FUNCTION_BLOCK Fase_Solida (* Fase solida (900): estocagem, alimentacao das prensas C-Press, polimero - HidrycoLib *)
  (* Standard: 61499-2 *)
  (* Version 1.5, 04/11/2026, Hidryco, Hidryco, 1.5: termica das bombas BO-900-01/02/03 NA (cfgTermicaNF = FALSE, campo: ligado = atuada). 1.4: velocidade de partida e PIDs das prensas em Hz (conversao no CLP). 1.3: pidCtl Pid1/2/3 com CycleTime 1000 ms (sem ele o calculo ciclico do pidSC ficava sem periodo). 1.2: sub-CATs Revezamento (horas por soprador, padrao do legado com o nome da elevatoria) e PID (ganho, integral, velocidade minima/maxima das 3 prensas). 1.0: fase solida (900, PCE LODO). Sub-CATs: LIT_900_01/02 (nivel dos tanques, 4-20 mA), FT_900_01/02/03/07 (vazao, comunicacao), SO_900_01/02, BO_900_01..03, BR_900_01/02 (Motor_Generico com ATV), VA_900_01/02, VB_900_03/04, VA_900_06..13 (Valvula_Coester on/off; VA_900_12 futura), AD_900_01..03 (Prensa_Vibropac; AD_900_03 futura), PP_900_01 (Preparador_Vibropac). Campo por symlink ${PATH}: djXXX (disjuntores do PCM LODO, XXX = equipamento), stsEmergenciaPainel (NF), stsMonitTrafo, stsMonitFonte, stsRemota1ComOk, stsRemota2Conexao (INT, connStatusInt); escrita cmdSV01/02/03/04/06/08 (solenoides, manual). *)
  PACKAGE Hidryco.HidrycoLib;
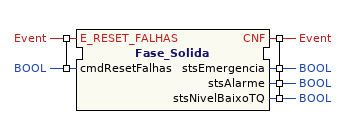
  EVENT_INPUT
    E_RESET_FALHAS WITH cmdResetFalhas; (* Reset pelo processo (fase solida e equipamentos) com cmdResetFalhas = TRUE *)
  END_EVENT
  EVENT_OUTPUT
    CNF WITH stsEmergencia, stsAlarme, stsNivelBaixoTQ; (* Status *)
  END_EVENT
  VAR_INPUT
    cmdResetFalhas : BOOL; (* TRUE = reset (com o evento E_RESET_FALHAS) *)
  END_VAR
  VAR_OUTPUT
    stsEmergencia : BOOL; (* Emergencia do PCM LODO *)
    stsAlarme : BOOL; (* Algum alarme da alimentacao/painel *)
    stsNivelBaixoTQ : BOOL; (* Tanques de estocagem em nivel baixo *)
  END_VAR
  FBS
    IThis : Fase_Solida_HMI(QI := TRUE);
    plcStart1 : plcStart(Prio := 10);
    Tick : E_CYCLE(DT := T#1s);
    Estocagem : basicEstocagemLodo;
    Alimentacao : basicAlimentacaoPrensas;
    Disjuntores1 : SYMLINKMULTIVARDST_854A896E88500D19(QI := TRUE, NAME1 := '$${PATH}djPCE', NAME2 := '$${PATH}djPCM', NAME3 := '$${PATH}djSO01', NAME4 := '$${PATH}djSO02', NAME5 := '$${PATH}djAD01', NAME6 := '$${PATH}djAD02', NAME7 := '$${PATH}djAD03', NAME8 := '$${PATH}djPP01', NAME9 := '$${PATH}djMN01', NAME10 := '$${PATH}djMN02', NAME11 := '$${PATH}djMN03', NAME12 := '$${PATH}djMN04', NAME13 := '$${PATH}djMN05', NAME14 := '$${PATH}djBO01', NAME15 := '$${PATH}djBO02', NAME16 := '$${PATH}djBO03'); {SET_ATTRIBUTE(Configuration.GenericFBType.InterfaceParams, Runtime.System#I:=16;VALUE${I$}:BOOL,BOOL,BOOL,BOOL,BOOL,BOOL,BOOL,BOOL,BOOL,BOOL,BOOL,BOOL,BOOL,BOOL,BOOL,BOOL)}
    Disjuntores2 : SYMLINKMULTIVARDST_854A896E88500D19(QI := TRUE, NAME1 := '$${PATH}djBR01', NAME2 := '$${PATH}djBR02', NAME3 := '$${PATH}djVA01', NAME4 := '$${PATH}djVA02', NAME5 := '$${PATH}djVE01', NAME6 := '$${PATH}djVE02', NAME7 := '$${PATH}djVA06', NAME8 := '$${PATH}djVA07', NAME9 := '$${PATH}djVA08', NAME10 := '$${PATH}djVA09', NAME11 := '$${PATH}djVA10', NAME12 := '$${PATH}djVA11', NAME13 := '$${PATH}djVA12', NAME14 := '$${PATH}djVA13', NAME15 := '$${PATH}djVB03', NAME16 := '$${PATH}djVB04'); {SET_ATTRIBUTE(Configuration.GenericFBType.InterfaceParams, Runtime.System#I:=16;VALUE${I$}:BOOL,BOOL,BOOL,BOOL,BOOL,BOOL,BOOL,BOOL,BOOL,BOOL,BOOL,BOOL,BOOL,BOOL,BOOL,BOOL)}
    Painel : SYMLINKMULTIVARDST_151ACB50A2F8223B2(QI := TRUE, NAME1 := '$${PATH}stsEmergenciaPainel', NAME2 := '$${PATH}stsMonitTrafo', NAME3 := '$${PATH}stsMonitFonte'); {SET_ATTRIBUTE(Configuration.GenericFBType.InterfaceParams, Runtime.System#I:=3;VALUE${I$}:BOOL,BOOL,BOOL)}
    Remota1 : SYMLINKMULTIVARDST_1559B0FF8170C9BA0(QI := TRUE, NAME1 := '$${PATH}stsRemota1ComOk'); {SET_ATTRIBUTE(Configuration.GenericFBType.InterfaceParams, Runtime.System#I:=1;VALUE${I$}:BOOL)}
    Remota2 : SYMLINKMULTIVARDST_5A03F112CD5D470(QI := TRUE, NAME1 := '$${PATH}stsRemota2Conexao'); {SET_ATTRIBUTE(Configuration.GenericFBType.InterfaceParams, Runtime.System#I:=1;VALUE${I$}:INT)}
    Solenoides1 : SYMLINKMULTIVARSRC_151ACB50A2F8223B2(QI := TRUE, NAME1 := '$${PATH}cmdSV01', NAME2 := '$${PATH}cmdSV02', NAME3 := '$${PATH}cmdSV03'); {SET_ATTRIBUTE(Configuration.GenericFBType.InterfaceParams, Runtime.System#I:=3;VALUE${I$}:BOOL,BOOL,BOOL)}
    Solenoides2 : SYMLINKMULTIVARSRC_151ACB50A2F8223B2(QI := TRUE, NAME1 := '$${PATH}cmdSV04', NAME2 := '$${PATH}cmdSV06', NAME3 := '$${PATH}cmdSV08'); {SET_ATTRIBUTE(Configuration.GenericFBType.InterfaceParams, Runtime.System#I:=3;VALUE${I$}:BOOL,BOOL,BOOL)}
    PersBO1 : PERSISTENCE_20652AC5DB8BA8AD5(QI := TRUE); {SET_ATTRIBUTE(Configuration.GenericFBType.InterfaceParams, Runtime.Standard#I:=3;input${I$}:UINT,UINT,UDINT)}
    PersBO2 : PERSISTENCE_20652AC5DB8BA8AD5(QI := TRUE); {SET_ATTRIBUTE(Configuration.GenericFBType.InterfaceParams, Runtime.Standard#I:=3;input${I$}:UINT,UINT,UDINT)}
    PersBO3 : PERSISTENCE_20652AC5DB8BA8AD5(QI := TRUE); {SET_ATTRIBUTE(Configuration.GenericFBType.InterfaceParams, Runtime.Standard#I:=3;input${I$}:UINT,UINT,UDINT)}
    Pid1 : pidCtl(CycleTime := 1000, Direction := TRUE, Bump := FALSE, ProhibitOutInc := FALSE, ProhibitOutDec := FALSE);
    Pid2 : pidCtl(CycleTime := 1000, Direction := TRUE, Bump := FALSE, ProhibitOutInc := FALSE, ProhibitOutDec := FALSE);
    Pid3 : pidCtl(CycleTime := 1000, Direction := TRUE, Bump := FALSE, ProhibitOutInc := FALSE, ProhibitOutDec := FALSE);
    LIT_900_01 : Sensor_Generico(pin_FC98F78ABCBC0A7E := TRUE, pin_CC8EEC06FF0C4430 := 'm', pin_6D3A2524C5D0F0D1 := 2);
    LIT_900_02 : Sensor_Generico(pin_FC98F78ABCBC0A7E := TRUE, pin_CC8EEC06FF0C4430 := 'm', pin_6D3A2524C5D0F0D1 := 2);
    FT_900_01 : Sensor_Generico(pin_D46B37D45FD5AF5D := TRUE, pin_0ECE7B3867B02E0B := TRUE, pin_CC8EEC06FF0C4430 := 'm3/h', pin_6D3A2524C5D0F0D1 := 1);
    FT_900_02 : Sensor_Generico(pin_D46B37D45FD5AF5D := TRUE, pin_0ECE7B3867B02E0B := TRUE, pin_CC8EEC06FF0C4430 := 'm3/h', pin_6D3A2524C5D0F0D1 := 1);
    FT_900_03 : Sensor_Generico(pin_D46B37D45FD5AF5D := TRUE, pin_0ECE7B3867B02E0B := TRUE, pin_CC8EEC06FF0C4430 := 'm3/h', pin_6D3A2524C5D0F0D1 := 1);
    FT_900_07 : Sensor_Generico(pin_D46B37D45FD5AF5D := TRUE, pin_0ECE7B3867B02E0B := TRUE, pin_CC8EEC06FF0C4430 := 'm3/h', pin_6D3A2524C5D0F0D1 := 1);
    SO_900_01 : Motor_Generico(pin_63EFEFB7C85EC93E := TRUE, pin_39489193B7758574 := 600.0);
    SO_900_02 : Motor_Generico(pin_63EFEFB7C85EC93E := TRUE, pin_39489193B7758574 := 600.0);
    BO_900_01 : Motor_Generico(pin_63EFEFB7C85EC93E := TRUE, pin_39489193B7758574 := 600.0, pin_66763E13F70A4420 := FALSE);
    BO_900_02 : Motor_Generico(pin_63EFEFB7C85EC93E := TRUE, pin_39489193B7758574 := 600.0, pin_66763E13F70A4420 := FALSE);
    BO_900_03 : Motor_Generico(pin_63EFEFB7C85EC93E := TRUE, pin_39489193B7758574 := 600.0, pin_66763E13F70A4420 := FALSE);
    BR_900_01 : Motor_Generico(pin_63EFEFB7C85EC93E := TRUE, pin_39489193B7758574 := 600.0);
    BR_900_02 : Motor_Generico(pin_63EFEFB7C85EC93E := TRUE, pin_39489193B7758574 := 600.0);
    VA_900_01 : Atuador_Coester;
    VA_900_02 : Atuador_Coester;
    VB_900_03 : Atuador_Coester;
    VB_900_04 : Atuador_Coester;
    VA_900_06 : Atuador_Coester;
    VA_900_07 : Atuador_Coester;
    VA_900_08 : Atuador_Coester;
    VA_900_09 : Atuador_Coester;
    VA_900_10 : Atuador_Coester;
    VA_900_11 : Atuador_Coester;
    VA_900_12 : Atuador_Coester(pin_FFAFC48D6FD3FF02 := FALSE);
    VA_900_13 : Atuador_Coester;
    AD_900_01 : Prensa_Vibropac;
    AD_900_02 : Prensa_Vibropac;
    AD_900_03 : Prensa_Vibropac(pin_FF2D8D14693482D2 := FALSE);
    PP_900_01 : Preparador_Vibropac;
    AlarmeSopradores : ALARM_BIT(TYPE := 1, ACKTYPE_1 := 2, ACTIVE := TRUE); {SET_ATTRIBUTE(HMI.AlarmText, Tanques de lodo: nenhum soprador disponível)}
    AlarmeNivelTQ : ALARM_BIT(TYPE := 1, ACKTYPE_1 := 2, ACTIVE := TRUE); {SET_ATTRIBUTE(HMI.AlarmText, Tanques de lodo: nível baixo - bombas suspensas)} {SET_ATTRIBUTE(HMI.AlarmClass, Warning)}
    AlarmeEmergencia : ALARM_BIT(TYPE := 1, ACKTYPE_1 := 2, ACTIVE := TRUE); {SET_ATTRIBUTE(HMI.AlarmText, PCM LODO: emergência acionada)}
    AlarmeRemota : ALARM_BIT(TYPE := 1, ACKTYPE_1 := 2, ACTIVE := TRUE); {SET_ATTRIBUTE(HMI.AlarmText, PCE LODO: remota sem comunicação)} {SET_ATTRIBUTE(HMI.AlarmClass, Warning)}
    AlarmeDisjuntor : ALARM_BIT(TYPE := 1, ACKTYPE_1 := 2, ACTIVE := TRUE); {SET_ATTRIBUTE(HMI.AlarmText, PCM LODO: disjuntor desligado)} {SET_ATTRIBUTE(HMI.AlarmClass, Warning)}
    AlarmeRota : ALARM_BIT(TYPE := 1, ACKTYPE_1 := 2, ACTIVE := TRUE); {SET_ATTRIBUTE(HMI.AlarmText, Alimentação das prensas: válvulas da rota não abriram)}
    AlarmeSemBomba : ALARM_BIT(TYPE := 1, ACKTYPE_1 := 2, ACTIVE := TRUE); {SET_ATTRIBUTE(HMI.AlarmText, Alimentação das prensas: sem bomba disponível)} {SET_ATTRIBUTE(HMI.AlarmClass, Warning)}
    AlarmeSemPartir : ALARM_BIT(TYPE := 1, ACKTYPE_1 := 2, ACTIVE := TRUE); {SET_ATTRIBUTE(HMI.AlarmText, Alimentação das prensas: prensa não partiu)} {SET_ATTRIBUTE(HMI.AlarmClass, Warning)}
    AlarmeFT : ALARM_BIT(TYPE := 1, ACKTYPE_1 := 2, ACTIVE := TRUE); {SET_ATTRIBUTE(HMI.AlarmText, Alimentação das prensas: medidor de vazão em falha)} {SET_ATTRIBUTE(HMI.AlarmClass, Warning)}
    Revezamento : Controle_Revezamento_2;
    PID : Controle_PID;
  END_FBS
  EVENT_CONNECTIONS
    plcStart1.FIRST_INIT TO IThis.F45AEED5C0881751;
    plcStart1.REDO_INIT TO IThis.F45AEED5C0881751;
    IThis.89CE2E9FA670B6C6 TO Disjuntores1.INIT;
    Disjuntores1.INITO TO Disjuntores2.INIT;
    Disjuntores2.INITO TO Painel.INIT;
    Painel.INITO TO Remota1.INIT;
    Remota1.INITO TO Remota2.INIT;
    Remota2.INITO TO Solenoides1.INIT;
    Solenoides1.INITO TO Solenoides2.INIT;
    Solenoides2.INITO TO Estocagem.243DC77CA0D0953F;
    Estocagem.5F76B62564497316 TO Alimentacao.13FEA6D5249A7B77;
    Alimentacao.8D3D86F80598A7BB TO IThis.AD1CFD9CF87E7BE8;
    Alimentacao.8D3D86F80598A7BB TO Tick.START;
    Alimentacao.8D3D86F80598A7BB TO PersBO1.INIT;
    PersBO1.INITO TO PersBO1.READ;
    PersBO1.READCNF TO Alimentacao.08CA7CB6A8F97690;
    Alimentacao.557985467D809489 TO PersBO1.WRITE;
    PersBO1.INITO TO PersBO2.INIT;
    PersBO2.INITO TO PersBO2.READ;
    PersBO2.READCNF TO Alimentacao.08CA7CB6A8F97690;
    Alimentacao.557985467D809489 TO PersBO2.WRITE;
    PersBO2.INITO TO PersBO3.INIT;
    PersBO3.INITO TO PersBO3.READ;
    PersBO3.READCNF TO Alimentacao.08CA7CB6A8F97690;
    Alimentacao.557985467D809489 TO PersBO3.WRITE;
    PersBO3.INITO TO AlarmeSopradores.INIT;
    AlarmeSopradores.INITO TO AlarmeSopradores.REQ_INITDATA;
    AlarmeSopradores.CNF_INITDATA TO AlarmeSopradores.ACTIVATE;
    AlarmeNivelTQ.INITO TO AlarmeNivelTQ.REQ_INITDATA;
    AlarmeNivelTQ.CNF_INITDATA TO AlarmeNivelTQ.ACTIVATE;
    AlarmeSopradores.INITO TO AlarmeNivelTQ.INIT;
    AlarmeEmergencia.INITO TO AlarmeEmergencia.REQ_INITDATA;
    AlarmeEmergencia.CNF_INITDATA TO AlarmeEmergencia.ACTIVATE;
    AlarmeNivelTQ.INITO TO AlarmeEmergencia.INIT;
    AlarmeRemota.INITO TO AlarmeRemota.REQ_INITDATA;
    AlarmeRemota.CNF_INITDATA TO AlarmeRemota.ACTIVATE;
    AlarmeEmergencia.INITO TO AlarmeRemota.INIT;
    AlarmeDisjuntor.INITO TO AlarmeDisjuntor.REQ_INITDATA;
    AlarmeDisjuntor.CNF_INITDATA TO AlarmeDisjuntor.ACTIVATE;
    AlarmeRemota.INITO TO AlarmeDisjuntor.INIT;
    AlarmeRota.INITO TO AlarmeRota.REQ_INITDATA;
    AlarmeRota.CNF_INITDATA TO AlarmeRota.ACTIVATE;
    AlarmeDisjuntor.INITO TO AlarmeRota.INIT;
    AlarmeSemBomba.INITO TO AlarmeSemBomba.REQ_INITDATA;
    AlarmeSemBomba.CNF_INITDATA TO AlarmeSemBomba.ACTIVATE;
    AlarmeRota.INITO TO AlarmeSemBomba.INIT;
    AlarmeSemPartir.INITO TO AlarmeSemPartir.REQ_INITDATA;
    AlarmeSemPartir.CNF_INITDATA TO AlarmeSemPartir.ACTIVATE;
    AlarmeSemBomba.INITO TO AlarmeSemPartir.INIT;
    AlarmeFT.INITO TO AlarmeFT.REQ_INITDATA;
    AlarmeFT.CNF_INITDATA TO AlarmeFT.ACTIVATE;
    AlarmeSemPartir.INITO TO AlarmeFT.INIT;
    AlarmeFT.INITO TO plcStart1.ACK_FIRST;
    Tick.EO TO Estocagem.E8C8FA9D941AAB25;
    Tick.EO TO Alimentacao.97FA92419A632264;
    Disjuntores1.CNF TO Alimentacao.856DAE0A3F3D97F7;
    Disjuntores2.CNF TO Alimentacao.856DAE0A3F3D97F7;
    Painel.CNF TO Alimentacao.19B51840153EBC5A;
    Remota1.CNF TO Alimentacao.939B3751BD07756D;
    Remota2.CNF TO Alimentacao.5748134B24BEF763;
    SO_900_01.9D4F26EE27EDF5B9 TO Estocagem.DFFA20E8FEFD328B;
    Estocagem.A37D04399243417C TO SO_900_01.21070E4B73BFECDC;
    SO_900_02.9D4F26EE27EDF5B9 TO Estocagem.DFFA20E8FEFD328B;
    Estocagem.A37D04399243417C TO SO_900_02.21070E4B73BFECDC;
    LIT_900_01.28A380156DB271B8 TO Estocagem.EA4444D55C79B643;
    LIT_900_02.28A380156DB271B8 TO Estocagem.EA4444D55C79B643;
    Alimentacao.8A05961272844DF6 TO Estocagem.EBAA94C91027AB04;
    Estocagem.820328527C60D44B TO VA_900_01.6AE7937B5439A162;
    Estocagem.820328527C60D44B TO VA_900_02.6AE7937B5439A162;
    Estocagem.820328527C60D44B TO VB_900_03.6AE7937B5439A162;
    Estocagem.820328527C60D44B TO VB_900_04.6AE7937B5439A162;
    Estocagem.DD4EDADF061294FF TO Alimentacao.CBCF1D50DEE68A86;
    AD_900_01.8111B44229D619D2 TO Alimentacao.38F5F6E182F651D4;
    Alimentacao.9C532436C7A3B461 TO AD_900_01.7E5F12997195C3C2;
    AD_900_02.8111B44229D619D2 TO Alimentacao.38F5F6E182F651D4;
    Alimentacao.9C532436C7A3B461 TO AD_900_02.7E5F12997195C3C2;
    AD_900_03.8111B44229D619D2 TO Alimentacao.38F5F6E182F651D4;
    Alimentacao.9C532436C7A3B461 TO AD_900_03.7E5F12997195C3C2;
    BO_900_01.9D4F26EE27EDF5B9 TO Alimentacao.CA246CEBE60B1023;
    Alimentacao.7490FED3332AEC1E TO BO_900_01.21070E4B73BFECDC;
    BO_900_02.9D4F26EE27EDF5B9 TO Alimentacao.CA246CEBE60B1023;
    Alimentacao.7490FED3332AEC1E TO BO_900_02.21070E4B73BFECDC;
    BO_900_03.9D4F26EE27EDF5B9 TO Alimentacao.CA246CEBE60B1023;
    Alimentacao.7490FED3332AEC1E TO BO_900_03.21070E4B73BFECDC;
    Alimentacao.7490FED3332AEC1E TO BR_900_01.21070E4B73BFECDC;
    Alimentacao.7490FED3332AEC1E TO BR_900_02.21070E4B73BFECDC;
    VA_900_06.CF6616D3CB5312F6 TO Alimentacao.6647071B86B2ADCE;
    Alimentacao.B985DE359C566AD4 TO VA_900_06.6AE7937B5439A162;
    VA_900_07.CF6616D3CB5312F6 TO Alimentacao.6647071B86B2ADCE;
    Alimentacao.B985DE359C566AD4 TO VA_900_07.6AE7937B5439A162;
    VA_900_08.CF6616D3CB5312F6 TO Alimentacao.6647071B86B2ADCE;
    Alimentacao.B985DE359C566AD4 TO VA_900_08.6AE7937B5439A162;
    VA_900_09.CF6616D3CB5312F6 TO Alimentacao.6647071B86B2ADCE;
    Alimentacao.B985DE359C566AD4 TO VA_900_09.6AE7937B5439A162;
    VA_900_10.CF6616D3CB5312F6 TO Alimentacao.6647071B86B2ADCE;
    Alimentacao.B985DE359C566AD4 TO VA_900_10.6AE7937B5439A162;
    VA_900_11.CF6616D3CB5312F6 TO Alimentacao.6647071B86B2ADCE;
    Alimentacao.B985DE359C566AD4 TO VA_900_11.6AE7937B5439A162;
    VA_900_12.CF6616D3CB5312F6 TO Alimentacao.6647071B86B2ADCE;
    Alimentacao.B985DE359C566AD4 TO VA_900_12.6AE7937B5439A162;
    VA_900_13.CF6616D3CB5312F6 TO Alimentacao.6647071B86B2ADCE;
    Alimentacao.B985DE359C566AD4 TO VA_900_13.6AE7937B5439A162;
    FT_900_01.28A380156DB271B8 TO Alimentacao.48ABB9D9BB2D6CEE;
    IThis.2286FBFA7E7E3034 TO Pid1.REQ_SP;
    FT_900_01.28A380156DB271B8 TO Pid1.REQ;
    Alimentacao.CF7635F428763261 TO Pid1.REQ;
    Pid1.CNF TO Alimentacao.37F5128277E33C7D;
    Pid1.C_CNF TO Alimentacao.37F5128277E33C7D;
    FT_900_02.28A380156DB271B8 TO Alimentacao.48ABB9D9BB2D6CEE;
    IThis.2286FBFA7E7E3034 TO Pid2.REQ_SP;
    FT_900_02.28A380156DB271B8 TO Pid2.REQ;
    Alimentacao.CF7635F428763261 TO Pid2.REQ;
    Pid2.CNF TO Alimentacao.37F5128277E33C7D;
    Pid2.C_CNF TO Alimentacao.37F5128277E33C7D;
    FT_900_03.28A380156DB271B8 TO Alimentacao.48ABB9D9BB2D6CEE;
    IThis.2286FBFA7E7E3034 TO Pid3.REQ_SP;
    FT_900_03.28A380156DB271B8 TO Pid3.REQ;
    Alimentacao.CF7635F428763261 TO Pid3.REQ;
    Pid3.CNF TO Alimentacao.37F5128277E33C7D;
    Pid3.C_CNF TO Alimentacao.37F5128277E33C7D;
    PP_900_01.0264E737EBBCA257 TO Alimentacao.2E29057D22A77FC3;
    Alimentacao.FAFF2EF1C05DA77F TO PP_900_01.8E41CA7EF16C6739;
    Alimentacao.F922E54EB08BF260 TO Solenoides1.REQ;
    Alimentacao.F922E54EB08BF260 TO Solenoides2.REQ;
    IThis.2286FBFA7E7E3034 TO Estocagem.C2DAB560DFFB8D5C;
    IThis.2286FBFA7E7E3034 TO Alimentacao.912D39602F9C91C5;
    IThis.94340A1957F06E33 TO Alimentacao.477B3CB066C0064B;
    IThis.DA6F3DD5304C4EDD TO Alimentacao.B672F1361E424ACE;
    IThis.EA322A066409681E TO Alimentacao.FBC24ECA7AD15CA0;
    Estocagem.12E6850BBBD0B68E TO IThis.0FDAAD8F71C680CA;
    Alimentacao.4D417ED96141B64B TO IThis.0FDAAD8F71C680CA;
    Estocagem.12E6850BBBD0B68E TO AlarmeSopradores.REQ;
    AlarmeSopradores.IND_1 TO IThis.0FDAAD8F71C680CA;
    IThis.EA322A066409681E TO AlarmeSopradores.ACK_C1;
    E_RESET_FALHAS TO AlarmeSopradores.ACK_C1;
    Estocagem.12E6850BBBD0B68E TO AlarmeNivelTQ.REQ;
    AlarmeNivelTQ.IND_1 TO IThis.0FDAAD8F71C680CA;
    IThis.EA322A066409681E TO AlarmeNivelTQ.ACK_C1;
    E_RESET_FALHAS TO AlarmeNivelTQ.ACK_C1;
    Alimentacao.4D417ED96141B64B TO AlarmeEmergencia.REQ;
    AlarmeEmergencia.IND_1 TO IThis.0FDAAD8F71C680CA;
    IThis.EA322A066409681E TO AlarmeEmergencia.ACK_C1;
    E_RESET_FALHAS TO AlarmeEmergencia.ACK_C1;
    Alimentacao.4D417ED96141B64B TO AlarmeRemota.REQ;
    AlarmeRemota.IND_1 TO IThis.0FDAAD8F71C680CA;
    IThis.EA322A066409681E TO AlarmeRemota.ACK_C1;
    E_RESET_FALHAS TO AlarmeRemota.ACK_C1;
    Alimentacao.4D417ED96141B64B TO AlarmeDisjuntor.REQ;
    AlarmeDisjuntor.IND_1 TO IThis.0FDAAD8F71C680CA;
    IThis.EA322A066409681E TO AlarmeDisjuntor.ACK_C1;
    E_RESET_FALHAS TO AlarmeDisjuntor.ACK_C1;
    Alimentacao.4D417ED96141B64B TO AlarmeRota.REQ;
    AlarmeRota.IND_1 TO IThis.0FDAAD8F71C680CA;
    IThis.EA322A066409681E TO AlarmeRota.ACK_C1;
    E_RESET_FALHAS TO AlarmeRota.ACK_C1;
    Alimentacao.4D417ED96141B64B TO AlarmeSemBomba.REQ;
    AlarmeSemBomba.IND_1 TO IThis.0FDAAD8F71C680CA;
    IThis.EA322A066409681E TO AlarmeSemBomba.ACK_C1;
    E_RESET_FALHAS TO AlarmeSemBomba.ACK_C1;
    Alimentacao.4D417ED96141B64B TO AlarmeSemPartir.REQ;
    AlarmeSemPartir.IND_1 TO IThis.0FDAAD8F71C680CA;
    IThis.EA322A066409681E TO AlarmeSemPartir.ACK_C1;
    E_RESET_FALHAS TO AlarmeSemPartir.ACK_C1;
    Alimentacao.4D417ED96141B64B TO AlarmeFT.REQ;
    AlarmeFT.IND_1 TO IThis.0FDAAD8F71C680CA;
    IThis.EA322A066409681E TO AlarmeFT.ACK_C1;
    E_RESET_FALHAS TO AlarmeFT.ACK_C1;
    E_RESET_FALHAS TO Alimentacao.E0DC297DC07DC5FB;
    E_RESET_FALHAS TO LIT_900_01.D21DAA5004F58516;
    E_RESET_FALHAS TO LIT_900_02.D21DAA5004F58516;
    E_RESET_FALHAS TO FT_900_01.D21DAA5004F58516;
    E_RESET_FALHAS TO FT_900_02.D21DAA5004F58516;
    E_RESET_FALHAS TO FT_900_03.D21DAA5004F58516;
    E_RESET_FALHAS TO FT_900_07.D21DAA5004F58516;
    E_RESET_FALHAS TO SO_900_01.BA30A65ADDA4ECC3;
    E_RESET_FALHAS TO SO_900_02.BA30A65ADDA4ECC3;
    E_RESET_FALHAS TO BO_900_01.BA30A65ADDA4ECC3;
    E_RESET_FALHAS TO BO_900_02.BA30A65ADDA4ECC3;
    E_RESET_FALHAS TO BO_900_03.BA30A65ADDA4ECC3;
    E_RESET_FALHAS TO BR_900_01.BA30A65ADDA4ECC3;
    E_RESET_FALHAS TO BR_900_02.BA30A65ADDA4ECC3;
    E_RESET_FALHAS TO VA_900_01.D903CD18EBE204D1;
    E_RESET_FALHAS TO VA_900_02.D903CD18EBE204D1;
    E_RESET_FALHAS TO VB_900_03.D903CD18EBE204D1;
    E_RESET_FALHAS TO VB_900_04.D903CD18EBE204D1;
    E_RESET_FALHAS TO VA_900_06.D903CD18EBE204D1;
    E_RESET_FALHAS TO VA_900_07.D903CD18EBE204D1;
    E_RESET_FALHAS TO VA_900_08.D903CD18EBE204D1;
    E_RESET_FALHAS TO VA_900_09.D903CD18EBE204D1;
    E_RESET_FALHAS TO VA_900_10.D903CD18EBE204D1;
    E_RESET_FALHAS TO VA_900_11.D903CD18EBE204D1;
    E_RESET_FALHAS TO VA_900_12.D903CD18EBE204D1;
    E_RESET_FALHAS TO VA_900_13.D903CD18EBE204D1;
    E_RESET_FALHAS TO AD_900_01.6BF17A43E520A528;
    E_RESET_FALHAS TO AD_900_02.6BF17A43E520A528;
    E_RESET_FALHAS TO AD_900_03.6BF17A43E520A528;
    E_RESET_FALHAS TO PP_900_01.92DC3CE3AA129B98;
    Alimentacao.8A05961272844DF6 TO CNF;
    Estocagem.DD4EDADF061294FF TO CNF;
    PID.75EB05A15DC6DC61 TO Pid1.REQ_PARA;
    PID.75EB05A15DC6DC61 TO Pid2.REQ_PARA;
    PID.75EB05A15DC6DC61 TO Pid3.REQ_PARA;
    Revezamento.62818F2F9E2138FC TO Estocagem.C2DAB560DFFB8D5C;
    Alimentacao.8D3D86F80598A7BB TO Revezamento.1DF068F97CBC55AD;
    Alimentacao.8D3D86F80598A7BB TO PID.117942CC3F34C94C;
    Estocagem.12E6850BBBD0B68E TO Revezamento.7D54AD64877107DE;
  END_CONNECTIONS
  DATA_CONNECTIONS
    PersBO1.output3 TO Alimentacao.B911BDD750DFDB18;
    Alimentacao.1115D73707983236 TO PersBO1.input3;
    PersBO2.output3 TO Alimentacao.0B46A3EB87E62664;
    Alimentacao.B5376FDD1F7B80EC TO PersBO2.input3;
    PersBO3.output3 TO Alimentacao.F9B917CCD98459B1;
    Alimentacao.4AE15F69ED84F18E TO PersBO3.input3;
    Disjuntores1.VALUE1 TO Alimentacao.4B9AB4FB6046D8EE;
    Disjuntores2.VALUE1 TO Alimentacao.1C7E6FC9EE536D0D;
    Disjuntores1.VALUE2 TO Alimentacao.F352CCB996881721;
    Disjuntores2.VALUE2 TO Alimentacao.B2F0010C50C459DF;
    Disjuntores1.VALUE3 TO Alimentacao.842E883449FD3557;
    Disjuntores2.VALUE3 TO Alimentacao.77D0D5AE9FA08670;
    Disjuntores1.VALUE4 TO Alimentacao.539AE49B193C0D44;
    Disjuntores2.VALUE4 TO Alimentacao.8E3376557963A36A;
    Disjuntores1.VALUE5 TO Alimentacao.299A09E7B67B47A1;
    Disjuntores2.VALUE5 TO Alimentacao.341C7D073810ED81;
    Disjuntores1.VALUE6 TO Alimentacao.F1AD4D08B9B3E19B;
    Disjuntores2.VALUE6 TO Alimentacao.9B9B7975525B3D51;
    Disjuntores1.VALUE7 TO Alimentacao.F9AFDD74B68569E8;
    Disjuntores2.VALUE7 TO Alimentacao.635621EAC24C7E9F;
    Disjuntores1.VALUE8 TO Alimentacao.A015D8C5AD7E44D6;
    Disjuntores2.VALUE8 TO Alimentacao.CFF227E520FF8AAB;
    Disjuntores1.VALUE9 TO Alimentacao.A2936012A1CB58B1;
    Disjuntores2.VALUE9 TO Alimentacao.B71059A1C4B0E360;
    Disjuntores1.VALUE10 TO Alimentacao.4FDDCD566D00E429;
    Disjuntores2.VALUE10 TO Alimentacao.7890B49E5275799F;
    Disjuntores1.VALUE11 TO Alimentacao.9F13912CAF6722CA;
    Disjuntores2.VALUE11 TO Alimentacao.651AFFD01F8F8841;
    Disjuntores1.VALUE12 TO Alimentacao.C0CD4D3BED37162D;
    Disjuntores2.VALUE12 TO Alimentacao.AA36A93C04F0663F;
    Disjuntores1.VALUE13 TO Alimentacao.F054F35A815A5F3B;
    Disjuntores2.VALUE13 TO Alimentacao.5365886519406CEA;
    Disjuntores1.VALUE14 TO Alimentacao.D38C2EC92076024C;
    Disjuntores2.VALUE14 TO Alimentacao.EBA41320B6D71E7A;
    Disjuntores1.VALUE15 TO Alimentacao.F3ED74F582F3070A;
    Disjuntores2.VALUE15 TO Alimentacao.1FB52CF6E301DAFF;
    Disjuntores1.VALUE16 TO Alimentacao.E8080276013928B8;
    Disjuntores2.VALUE16 TO Alimentacao.0C6B46DC80495D9D;
    Painel.VALUE1 TO Alimentacao.DE87224B5A8EF166;
    Painel.VALUE2 TO Alimentacao.554D2A3603C18677;
    Painel.VALUE3 TO Alimentacao.DFA71CBA2E1C52C4;
    Remota1.VALUE1 TO Alimentacao.82720E0D992C7F0F;
    Remota2.VALUE1 TO Alimentacao.9252FB36847BBAB8;
    SO_900_01.EBDC9E59C4286586 TO Estocagem.9D0A018985052F58;
    SO_900_01.40A5976BFB296133 TO Estocagem.C050A723D1972718;
    Estocagem.6EEF3183DA620253 TO SO_900_01.87DAE15414E7C412;
    Estocagem.821D8F0728BFD8D2 TO SO_900_01.85953C7B9294A9BF;
    SO_900_02.EBDC9E59C4286586 TO Estocagem.6442D6171574AD0F;
    SO_900_02.40A5976BFB296133 TO Estocagem.DB889EF87AAB0D82;
    Estocagem.8F8F344FCE172148 TO SO_900_02.87DAE15414E7C412;
    Estocagem.821D8F0728BFD8D2 TO SO_900_02.85953C7B9294A9BF;
    LIT_900_01.E6F78A591442B69F TO Estocagem.76186D6114386881;
    LIT_900_01.726640D1704B3F86 TO Estocagem.DEE813645F20FA9B;
    LIT_900_02.E6F78A591442B69F TO Estocagem.8747D35EC434F184;
    LIT_900_02.726640D1704B3F86 TO Estocagem.284C3EA5513A6D62;
    Alimentacao.1322393E4B988CAC TO Estocagem.8603BC9EB66FE144;
    Estocagem.937510DD507F2D1B TO VA_900_01.05903B4B679AA14E;
    Estocagem.937510DD507F2D1B TO VA_900_02.05903B4B679AA14E;
    Estocagem.937510DD507F2D1B TO VB_900_03.05903B4B679AA14E;
    Estocagem.937510DD507F2D1B TO VB_900_04.05903B4B679AA14E;
    Estocagem.9185345097862782 TO Alimentacao.70D9A60B95DEEE36;
    AD_900_01.D0AE1B8C5839DEE7 TO Alimentacao.65110DE39233F1DF;
    AD_900_01.4BC1097F03D3F72F TO Alimentacao.F2B23EF191CE5815;
    AD_900_01.984D9CCB4CB171BC TO Alimentacao.EA7AE03BB2089BBC;
    Alimentacao.61DAE1163D383245 TO AD_900_01.12D984BF9E1FDA1E;
    AD_900_02.D0AE1B8C5839DEE7 TO Alimentacao.77FAB1BD40DD3B80;
    AD_900_02.4BC1097F03D3F72F TO Alimentacao.841BFE40D529C6D2;
    AD_900_02.984D9CCB4CB171BC TO Alimentacao.04A6E0D53C4D9443;
    Alimentacao.7BECFC93E64F7C4C TO AD_900_02.12D984BF9E1FDA1E;
    AD_900_03.D0AE1B8C5839DEE7 TO Alimentacao.274510EEDF09C6C1;
    AD_900_03.4BC1097F03D3F72F TO Alimentacao.6BCEE4FB5283E200;
    AD_900_03.984D9CCB4CB171BC TO Alimentacao.4EEBC2ED0DBBF0E1;
    Alimentacao.0886EC6A983E53EF TO AD_900_03.12D984BF9E1FDA1E;
    BO_900_01.EBDC9E59C4286586 TO Alimentacao.948786DC7FA5A6CE;
    BO_900_01.40A5976BFB296133 TO Alimentacao.7764C36D58E005D1;
    BO_900_01.C5DF7BA69D90B1CF TO Alimentacao.83CDCBFE9DEDD3FA;
    Alimentacao.3D555F8584F77E3E TO BO_900_01.87DAE15414E7C412;
    Alimentacao.539E2B4F1B6EB82B TO BO_900_01.F94ABA993E8E9FF4;
    Alimentacao.37F7D293861FDD8C TO BO_900_01.85953C7B9294A9BF;
    BO_900_02.EBDC9E59C4286586 TO Alimentacao.B7E8FF7BEBB89AF3;
    BO_900_02.40A5976BFB296133 TO Alimentacao.41C84D6CB5F8D848;
    BO_900_02.C5DF7BA69D90B1CF TO Alimentacao.1A1D9754A8468CF5;
    Alimentacao.BF55FDEF007D89FD TO BO_900_02.87DAE15414E7C412;
    Alimentacao.F2E13B217536BA96 TO BO_900_02.F94ABA993E8E9FF4;
    Alimentacao.37F7D293861FDD8C TO BO_900_02.85953C7B9294A9BF;
    BO_900_03.EBDC9E59C4286586 TO Alimentacao.5A6232E8B7292CDD;
    BO_900_03.40A5976BFB296133 TO Alimentacao.32464E571E89C87D;
    BO_900_03.C5DF7BA69D90B1CF TO Alimentacao.BE30680B6785F53B;
    Alimentacao.15B6EA39D5978533 TO BO_900_03.87DAE15414E7C412;
    Alimentacao.3A30521D5984EF99 TO BO_900_03.F94ABA993E8E9FF4;
    Alimentacao.37F7D293861FDD8C TO BO_900_03.85953C7B9294A9BF;
    Alimentacao.37F7D293861FDD8C TO BR_900_01.85953C7B9294A9BF;
    Alimentacao.37F7D293861FDD8C TO BR_900_02.85953C7B9294A9BF;
    VA_900_06.5EDB2238B0F9A6B6 TO Alimentacao.EAEBC6AA04FEFCE7;
    VA_900_06.C1396A09200C7A2F TO Alimentacao.0160D0A62EA49008;
    VA_900_06.904DD3246D8E0F2F TO Alimentacao.4DCA85ED8ED727AC;
    Alimentacao.09388B5323AA3765 TO VA_900_06.05903B4B679AA14E;
    Alimentacao.A7CB426F9568B620 TO VA_900_06.DD850CDC4ADBDD2B;
    VA_900_07.5EDB2238B0F9A6B6 TO Alimentacao.260161B67AA60DC8;
    VA_900_07.C1396A09200C7A2F TO Alimentacao.78E29B18EA62877A;
    VA_900_07.904DD3246D8E0F2F TO Alimentacao.4F349E1228AFA18C;
    Alimentacao.AD2094C9498D759A TO VA_900_07.05903B4B679AA14E;
    Alimentacao.85D68BAB1621B6ED TO VA_900_07.DD850CDC4ADBDD2B;
    VA_900_08.5EDB2238B0F9A6B6 TO Alimentacao.5D2228E3EC8A6E1D;
    VA_900_08.C1396A09200C7A2F TO Alimentacao.E7A0AAF9B673D116;
    VA_900_08.904DD3246D8E0F2F TO Alimentacao.F47AE21FE590F0B3;
    Alimentacao.0A83E200DBF274DA TO VA_900_08.05903B4B679AA14E;
    Alimentacao.D72F280458923969 TO VA_900_08.DD850CDC4ADBDD2B;
    VA_900_09.5EDB2238B0F9A6B6 TO Alimentacao.AFE22666313FA87F;
    VA_900_09.C1396A09200C7A2F TO Alimentacao.656542BCD835F282;
    VA_900_09.904DD3246D8E0F2F TO Alimentacao.C008B33DFC39701B;
    Alimentacao.64C7E137F02EE9D7 TO VA_900_09.05903B4B679AA14E;
    Alimentacao.77D4E686879E7239 TO VA_900_09.DD850CDC4ADBDD2B;
    VA_900_10.5EDB2238B0F9A6B6 TO Alimentacao.37E7DA5192455D76;
    VA_900_10.C1396A09200C7A2F TO Alimentacao.706657C3D65F7F40;
    VA_900_10.904DD3246D8E0F2F TO Alimentacao.CC429EBE88373900;
    Alimentacao.1196AAA785140AD5 TO VA_900_10.05903B4B679AA14E;
    Alimentacao.85FEEEECD707E5BA TO VA_900_10.DD850CDC4ADBDD2B;
    VA_900_11.5EDB2238B0F9A6B6 TO Alimentacao.BDD83839263E31A1;
    VA_900_11.C1396A09200C7A2F TO Alimentacao.0BF81BEEF6EED279;
    VA_900_11.904DD3246D8E0F2F TO Alimentacao.58D7F1A138120A11;
    Alimentacao.11B4927E17D401ED TO VA_900_11.05903B4B679AA14E;
    Alimentacao.60F03D282CD92FBF TO VA_900_11.DD850CDC4ADBDD2B;
    VA_900_12.5EDB2238B0F9A6B6 TO Alimentacao.0EB99790809C97DD;
    VA_900_12.C1396A09200C7A2F TO Alimentacao.85DCC3F2A49D036D;
    VA_900_12.904DD3246D8E0F2F TO Alimentacao.E64E50A12946C6F7;
    Alimentacao.EDCFAA44360A7A3E TO VA_900_12.05903B4B679AA14E;
    Alimentacao.2CA326C6E7119016 TO VA_900_12.DD850CDC4ADBDD2B;
    VA_900_13.5EDB2238B0F9A6B6 TO Alimentacao.1265105CC55986A5;
    VA_900_13.C1396A09200C7A2F TO Alimentacao.034CCB38CD43E88F;
    VA_900_13.904DD3246D8E0F2F TO Alimentacao.4BD9CB54C9563BCC;
    Alimentacao.AA673A290EB62EF4 TO VA_900_13.05903B4B679AA14E;
    Alimentacao.DB9D8913794AE690 TO VA_900_13.DD850CDC4ADBDD2B;
    FT_900_01.D7422D307E6AF52D TO Alimentacao.E11687C0F6E4D8D0;
    FT_900_01.726640D1704B3F86 TO Alimentacao.34CF43065C440B3F;
    FT_900_01.D7422D307E6AF52D TO Pid1.Pv;
    IThis.49434B52BAD72F2D TO Pid1.Sp;
    Alimentacao.AC7C96EC320F9B56 TO Pid1.Mode;
    Alimentacao.66CC0FC8380DE7A9 TO Pid1.PresetValue;
    Pid1.Out TO Alimentacao.EF0418ED47F514A0;
    FT_900_02.D7422D307E6AF52D TO Alimentacao.0B775DA830BA5C8F;
    FT_900_02.726640D1704B3F86 TO Alimentacao.BF4060DB062B029B;
    FT_900_02.D7422D307E6AF52D TO Pid2.Pv;
    IThis.76E9ED00F32CFE6B TO Pid2.Sp;
    Alimentacao.8D0D9C2E90DCA136 TO Pid2.Mode;
    Alimentacao.82217E0576C4A321 TO Pid2.PresetValue;
    Pid2.Out TO Alimentacao.CB7E7E5A60558086;
    FT_900_03.D7422D307E6AF52D TO Alimentacao.1C872E508B6F9CCA;
    FT_900_03.726640D1704B3F86 TO Alimentacao.6DEAF5F9074BEFF6;
    FT_900_03.D7422D307E6AF52D TO Pid3.Pv;
    IThis.9A1935965FF11A1D TO Pid3.Sp;
    Alimentacao.580E8B452F14C837 TO Pid3.Mode;
    Alimentacao.F7E26881AF4B195B TO Pid3.PresetValue;
    Pid3.Out TO Alimentacao.0398A48B9177A287;
    PP_900_01.5924057DB679FD7F TO Alimentacao.F50C4FB10C56E01C;
    PP_900_01.1330DA43C77FB0EB TO Alimentacao.1B803ED11E2532F9;
    PP_900_01.278FA7DE98B71B84 TO Alimentacao.CC53CD434F3E136E;
    Alimentacao.CE3A2F0FFB2A4E6D TO PP_900_01.DB86CBF02B2705F4;
    Alimentacao.60CC14D8DBDCF308 TO Solenoides1.VALUE1;
    Alimentacao.253C46304686EE40 TO Solenoides1.VALUE2;
    Alimentacao.9AE50630E8A856E9 TO Solenoides1.VALUE3;
    Alimentacao.28A4416677CA3C6A TO Solenoides2.VALUE1;
    Alimentacao.21FE5B252B52D38C TO Solenoides2.VALUE2;
    Alimentacao.2A1E389F770A9C7F TO Solenoides2.VALUE3;
    IThis.75C48C19F662F275 TO Estocagem.5CF5D34DC0BD4690;
    IThis.22AD5AC875BC0F3A TO Estocagem.834BCC8A73E45242;
    IThis.1683EE138AB36942 TO Estocagem.6A41927EA4F7A44E;
    IThis.49434B52BAD72F2D TO Alimentacao.831130D22BEBE078;
    IThis.76E9ED00F32CFE6B TO Alimentacao.CF86D1D755F0EA89;
    IThis.9A1935965FF11A1D TO Alimentacao.35630ED20F729613;
    IThis.C5C888AF0BB9838A TO Alimentacao.3CE89723CC83D95B;
    IThis.EC8188235095061D TO Alimentacao.C297DFFBB305E08D;
    IThis.BB8CB73AEC41AFB6 TO Alimentacao.6540F6059C1CADFB;
    IThis.852A633C619D78DF TO Alimentacao.0F2A42F20BB3A299;
    IThis.7AEF88FD51FDF12B TO Alimentacao.6EADB4D7BECA8D09;
    IThis.6BD2979D7880F624 TO Alimentacao.01D9A373E0929133;
    IThis.14A916BBB29783A2 TO Alimentacao.AA3E9DEF7B14FC07;
    IThis.C1D7E1AD99B844D5 TO Alimentacao.90A8AB90CFE56298;
    IThis.4B9E3E283F7B0C32 TO Alimentacao.052CCF025B5CF1E6;
    IThis.827B894171AEFAE0 TO Alimentacao.AEE5CBA91FD7B8C0;
    IThis.CC007DD46872FCB9 TO Alimentacao.92496204688A25B6;
    IThis.07EAED9390EBE189 TO Alimentacao.9B16B5CD8598F0FE;
    IThis.E5D36800A163DA06 TO Alimentacao.E768577E71FC29DC;
    IThis.9436C2F5462D6C4B TO Alimentacao.287E3CB21FEE06B9;
    IThis.09360E0486758B0D TO Alimentacao.9F60FEAA00C8DAD0;
    IThis.5006944B41B9FF77 TO Alimentacao.4FC52CF361E2E60C;
    Estocagem.0C2557554843B422 TO IThis.110B7745F6B54438;
    Estocagem.0C18C6251210ADD2 TO IThis.A95EFB2487615573;
    Estocagem.4235B19D4DDCC680 TO IThis.D4D97E1ACC759832;
    Estocagem.00131AAE1783E6A4 TO IThis.20AD366CDD94A9A3;
    Estocagem.27E22A4C9A4D8B67 TO IThis.B26669A5A84C4CC7;
    Estocagem.9185345097862782 TO IThis.9E5208DD14F5BD28;
    Estocagem.7A648FEA2F2E214A TO IThis.FF8604009D2A1731;
    Alimentacao.D719943085A661DC TO IThis.FD33BA674F199A2D;
    Alimentacao.7ABDDDB4AC047B40 TO IThis.47F04DE0966781D0;
    Alimentacao.EEF5EE0476E38158 TO IThis.DCEDC83B6145E7B1;
    Alimentacao.1C58EC4E4D6007CF TO IThis.EC6741C22B920EC4;
    Alimentacao.3B3BA86239824893 TO IThis.44EA220F7CB20FE3;
    Alimentacao.3668184FE0033268 TO IThis.C4038C90B52ACFF2;
    Alimentacao.8CDFD98CD3EFB259 TO IThis.A57197B6D74E3F3A;
    Alimentacao.8C2711D878B9AC5E TO IThis.3123A4CB92CAF55B;
    Alimentacao.BB3E6BCFC6AF1E38 TO IThis.772561770269900E;
    Alimentacao.DF31C371889E2274 TO IThis.398054DBC899C47E;
    Alimentacao.16341BB29A3C6F44 TO IThis.ED2141003596C6A0;
    Alimentacao.E71239536EFCF901 TO IThis.6FAF687D8B3E3E9C;
    Alimentacao.FBFF69BE7DE7E92A TO IThis.C739ADEA6D3C2837;
    Alimentacao.DABC56E6789EBDFB TO IThis.EE7172649A5770B4;
    Alimentacao.75E3B37E3578B9B2 TO IThis.5C3A4EBB1F23E5E7;
    Alimentacao.3A28F1E50DEF39F0 TO IThis.CC2D4B57EABA4F30;
    Alimentacao.EDE63BC2D534A388 TO IThis.43D2A3DA6B492647;
    Alimentacao.A6216B2CB75B6248 TO IThis.1D125FF4D75E807F;
    Alimentacao.DCFBAD76FD6DAC8A TO IThis.0FDFA1687EBDF6BB;
    Alimentacao.F44FD4A3D46566D4 TO IThis.9732E39322BDC91F;
    Alimentacao.E8F08415D1DE11AE TO IThis.19E815567D1C0103;
    Alimentacao.153BDE356C7E9BEA TO IThis.3E595E18CED9210D;
    Alimentacao.28634CDA5A89EA26 TO IThis.5E77C597D0181EFB;
    Alimentacao.57C5F71A067DD1B0 TO IThis.649160467445F4D8;
    Alimentacao.7932648D00F8B909 TO IThis.BD281849B3805537;
    Alimentacao.F378C93E70C9BC6C TO IThis.E34FF4D515E91AA3;
    Alimentacao.1322393E4B988CAC TO IThis.609B7773C5AA9D8D;
    Alimentacao.F6BBD672B702660F TO IThis.48DDFF06CB0DB57A;
    Alimentacao.B7F2CA425EC4E9E5 TO IThis.26A723406833679C;
    Alimentacao.4CFE0F5C97B9A171 TO IThis.DC8DEE0357A69788;
    Alimentacao.0BA3DFBF7BC917B6 TO IThis.E4B031F6683EC293;
    Alimentacao.DD0E1AA5D8A1DB26 TO IThis.012A50662A7C6CA6;
    Alimentacao.42975C96291AF6C2 TO IThis.2156A1525B988227;
    Alimentacao.5C804F1F7A91C337 TO IThis.A97E1235B4E4F47D;
    Alimentacao.59CAA41FF7F076C8 TO IThis.FE42C17BA14CFDF9;
    Alimentacao.D7727D91DD4BF548 TO IThis.6D5990A0ACA9F64C;
    Alimentacao.BEDB08F04967A6AF TO IThis.3B2E83E1E2181023;
    Alimentacao.712DA676390F489B TO IThis.282F57890E4910EA;
    Alimentacao.3EAEFAB9CF3845DF TO IThis.186FE869732C3A93;
    Alimentacao.81F88C6586FE748B TO IThis.D9D46ED2B3C829B1;
    Alimentacao.01F97979450409F0 TO IThis.3E23612E665F8916;
    Alimentacao.192257EE9070D8F5 TO IThis.9D6FF92E38B824A4;
    Estocagem.00131AAE1783E6A4 TO AlarmeSopradores.INP;
    AlarmeSopradores.STATE_1 TO IThis.D610D1C2A453F4AC;
    Estocagem.9185345097862782 TO AlarmeNivelTQ.INP;
    AlarmeNivelTQ.STATE_1 TO IThis.D2EA6A26C7F1B9D2;
    Alimentacao.1322393E4B988CAC TO AlarmeEmergencia.INP;
    AlarmeEmergencia.STATE_1 TO IThis.117470FCC1C36006;
    Alimentacao.4CFE0F5C97B9A171 TO AlarmeRemota.INP;
    AlarmeRemota.STATE_1 TO IThis.9239655AC6655482;
    Alimentacao.59CAA41FF7F076C8 TO AlarmeDisjuntor.INP;
    AlarmeDisjuntor.STATE_1 TO IThis.87E1350DB3E51FD0;
    Alimentacao.BEDB08F04967A6AF TO AlarmeRota.INP;
    AlarmeRota.STATE_1 TO IThis.0A46A1A5475DFF34;
    Alimentacao.D7727D91DD4BF548 TO AlarmeSemBomba.INP;
    AlarmeSemBomba.STATE_1 TO IThis.48D0207A23D83E95;
    Alimentacao.712DA676390F489B TO AlarmeSemPartir.INP;
    AlarmeSemPartir.STATE_1 TO IThis.802A5CD9C94AA734;
    Alimentacao.3EAEFAB9CF3845DF TO AlarmeFT.INP;
    AlarmeFT.STATE_1 TO IThis.C8DD695DFF1FA11F;
    cmdResetFalhas TO Alimentacao.3DBC80F4FE0835E7;
    cmdResetFalhas TO LIT_900_01.1908F43CB878F5E7;
    cmdResetFalhas TO LIT_900_02.1908F43CB878F5E7;
    cmdResetFalhas TO FT_900_01.1908F43CB878F5E7;
    cmdResetFalhas TO FT_900_02.1908F43CB878F5E7;
    cmdResetFalhas TO FT_900_03.1908F43CB878F5E7;
    cmdResetFalhas TO FT_900_07.1908F43CB878F5E7;
    cmdResetFalhas TO SO_900_01.C2F1E9C0FB076F17;
    cmdResetFalhas TO SO_900_02.C2F1E9C0FB076F17;
    cmdResetFalhas TO BO_900_01.C2F1E9C0FB076F17;
    cmdResetFalhas TO BO_900_02.C2F1E9C0FB076F17;
    cmdResetFalhas TO BO_900_03.C2F1E9C0FB076F17;
    cmdResetFalhas TO BR_900_01.C2F1E9C0FB076F17;
    cmdResetFalhas TO BR_900_02.C2F1E9C0FB076F17;
    cmdResetFalhas TO VA_900_01.C82CBBE25FC56079;
    cmdResetFalhas TO VA_900_02.C82CBBE25FC56079;
    cmdResetFalhas TO VB_900_03.C82CBBE25FC56079;
    cmdResetFalhas TO VB_900_04.C82CBBE25FC56079;
    cmdResetFalhas TO VA_900_06.C82CBBE25FC56079;
    cmdResetFalhas TO VA_900_07.C82CBBE25FC56079;
    cmdResetFalhas TO VA_900_08.C82CBBE25FC56079;
    cmdResetFalhas TO VA_900_09.C82CBBE25FC56079;
    cmdResetFalhas TO VA_900_10.C82CBBE25FC56079;
    cmdResetFalhas TO VA_900_11.C82CBBE25FC56079;
    cmdResetFalhas TO VA_900_12.C82CBBE25FC56079;
    cmdResetFalhas TO VA_900_13.C82CBBE25FC56079;
    cmdResetFalhas TO AD_900_01.38D2DBD6E8AAFA91;
    cmdResetFalhas TO AD_900_02.38D2DBD6E8AAFA91;
    cmdResetFalhas TO AD_900_03.38D2DBD6E8AAFA91;
    cmdResetFalhas TO PP_900_01.1C1DE110A3771399;
    Alimentacao.1322393E4B988CAC TO stsEmergencia;
    Alimentacao.192257EE9070D8F5 TO stsAlarme;
    Estocagem.9185345097862782 TO stsNivelBaixoTQ;
    PID.4F45CBCE24FA8775 TO Pid1.Gain;
    PID.5D86C7647B367BF7 TO Pid1.IntegralTime;
    PID.8B11A5B11AA557C3 TO Pid1.OutMin;
    PID.E7AF90225A9267BD TO Pid1.OutMax;
    PID.4F45CBCE24FA8775 TO Pid2.Gain;
    PID.5D86C7647B367BF7 TO Pid2.IntegralTime;
    PID.8B11A5B11AA557C3 TO Pid2.OutMin;
    PID.E7AF90225A9267BD TO Pid2.OutMax;
    PID.4F45CBCE24FA8775 TO Pid3.Gain;
    PID.5D86C7647B367BF7 TO Pid3.IntegralTime;
    PID.8B11A5B11AA557C3 TO Pid3.OutMin;
    PID.E7AF90225A9267BD TO Pid3.OutMax;
    Revezamento.E20C11B2DD910C9B TO Estocagem.7307922C026394A4;
    Revezamento.8F7C57B973CE6721 TO Estocagem.ABC6D729A9607229;
    Revezamento.B121C963D16B0207 TO Estocagem.F2FB54ACA0B1231D;
    Estocagem.C56DE563E1383C2E TO Revezamento.BCDE1E145B7C7428;
    Estocagem.6097DB009BDB40DE TO Revezamento.B99EA94F80E94BD2;
    Estocagem.53980AC2D919D417 TO Revezamento.30C56EFD8B8A4EB9;
  END_CONNECTIONS
END_FUNCTION_BLOCK
